ABB RAPID module: Weld1.mod

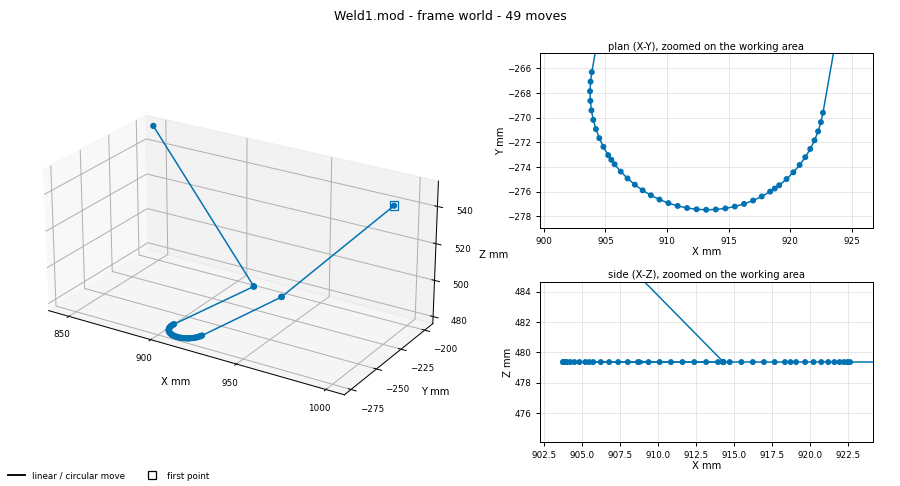
[picture p0: tool path of Weld1.mod in frame world, 49 of 50 moves have a stored position in this frame; points joined in program order, loops and branches not executed]
%%%
  VERSION:1
  LANGUAGE:ENGLISH
%%%
MODULE MOD_Weld1

    ! -------------------------------
    ! Define customized variables here
    ! ...

	! Tool variables:
	PERS tooldata Weldgun := [TRUE,[[-4.000,0.000,371.300],[0.92387953,0.00000000,0.38268343,0.00000001]],[1,[0,0,20],[1,0,0,0],0,0,0.005]];

	! Reference variables:
	PERS wobjdata WeldingReference := [FALSE, TRUE, "", [[0,0,0],[1,0,0,0]],[[907.213,-302.346,276.168],[0.70442562,0.70442562,-0.06151869,-0.06151869]]];

	PROC Main()
		ConfJ \On;
		ConfL \Off;
		! Program generated by VerticalBot Studio for ABB IRB 2600-12/1.65 on 25/10/2026 12:00:00
		! Using nominal kinematics.
		! show Weld gun
		MoveAbsJ [[-12.555800,6.650190,11.177100,0.026927,72.173900,-2.607590],[9E+09,9E+09,9E+09,9E+09,9E+09,9E+09]],v1000,z1,Weldgun \WObj:=WeldingReference;
		SetRPM 70.0;
		MoveL [[80.178,273.912,-94.776],[0.27080492,-0.27039115,-0.65336714,0.65319576],[-1,0,-1,0],[9E+09,9E+09,9E+09,9E+09,9E+09,9E+09]],[16.67,500,5000,1000],z1,Weldgun \WObj:=WeldingReference;
		MoveL [[9.468,203.201,-94.776],[0.27080492,-0.27039115,-0.65336714,0.65319576],[-1,0,-1,0],[9E+09,9E+09,9E+09,9E+09,9E+09,9E+09]],[16.67,500,5000,1000],z1,Weldgun \WObj:=WeldingReference;
		GunOn;
		MoveL [[9.468,203.201,-94.776],[0.27080492,-0.27039115,-0.65336714,0.65319576],[-1,0,-1,0],[9E+09,9E+09,9E+09,9E+09,9E+09,9E+09]],[16.67,500,5000,1000],z1,Weldgun \WObj:=WeldingReference;
		MoveL [[9.521,203.201,-94.770],[0.27059813,-0.27059797,-0.65328151,0.65328145],[-1,0,-1,0],[9E+09,9E+09,9E+09,9E+09,9E+09,9E+09]],[16.67,500,5000,1000],z1,Weldgun \WObj:=WeldingReference;
		MoveL [[9.521,203.201,-34.925],[0.26109596,-0.28004323,-0.64928868,0.65713689],[-1,-1,-1,0],[9E+09,9E+09,9E+09,9E+09,9E+09,9E+09]],[16.67,500,5000,1000],z1,Weldgun \WObj:=WeldingReference;
		MoveL [[9.489,203.201,-34.145],[0.23425026,-0.30675221,-0.65944853,0.64510273],[-1,-1,0,0],[9E+09,9E+09,9E+09,9E+09,9E+09,9E+09]],[16.67,500,5000,1000],z1,Weldgun \WObj:=WeldingReference;
		MoveL [[9.394,203.201,-33.370],[0.20701375,-0.33294335,-0.66849979,0.63198265],[-1,-1,0,0],[9E+09,9E+09,9E+09,9E+09,9E+09,9E+09]],[16.67,500,5000,1000],z1,Weldgun \WObj:=WeldingReference;
		MoveL [[9.235,203.201,-32.605],[0.17943264,-0.35858122,-0.67642029,0.61780177],[-1,-1,0,0],[9E+09,9E+09,9E+09,9E+09,9E+09,9E+09]],[16.67,500,5000,1000],z1,Weldgun \WObj:=WeldingReference;
		MoveL [[9.014,203.201,-31.857],[0.15154219,-0.38361099,-0.68321444,0.60257415],[-1,-1,0,0],[9E+09,9E+09,9E+09,9E+09,9E+09,9E+09]],[16.67,500,5000,1000],z1,Weldgun \WObj:=WeldingReference;
		MoveL [[8.732,203.201,-31.128],[0.12340353,-0.40798899,-0.68885701,0.58633828],[-1,-1,0,0],[9E+09,9E+09,9E+09,9E+09,9E+09,9E+09]],[16.67,500,5000,1000],z1,Weldgun \WObj:=WeldingReference;
		MoveL [[8.391,203.201,-30.426],[0.09505233,-0.43169103,-0.69333556,0.56911660],[-1,-1,0,0],[9E+09,9E+09,9E+09,9E+09,9E+09,9E+09]],[16.67,500,5000,1000],z1,Weldgun \WObj:=WeldingReference;
		MoveL [[7.994,203.201,-29.753],[0.06655006,-0.45466761,-0.69664493,0.55093947],[-1,-1,0,0],[9E+09,9E+09,9E+09,9E+09,9E+09,9E+09]],[16.67,500,5000,1000],z1,Weldgun \WObj:=WeldingReference;
		MoveL [[7.544,203.201,-29.116],[0.03792629,-0.47687790,-0.69878733,0.53183205],[-1,-1,0,0],[9E+09,9E+09,9E+09,9E+09,9E+09,9E+09]],[16.67,500,5000,1000],z1,Weldgun \WObj:=WeldingReference;
		MoveL [[7.042,203.201,-28.517],[0.01240330,-0.49395227,-0.70281556,0.51176909],[-1,-1,0,0],[9E+09,9E+09,9E+09,9E+09,9E+09,9E+09]],[16.67,500,5000,1000],z1,Weldgun \WObj:=WeldingReference;
		MoveL [[6.733,203.201,-28.192],[0.00416831,0.50587340,0.70291668,-0.49998286],[-1,-1,0,0],[9E+09,9E+09,9E+09,9E+09,9E+09,9E+09]],[16.67,500,5000,1000],z1,Weldgun \WObj:=WeldingReference;
		MoveL [[6.408,203.201,-27.883],[0.02374061,0.52184249,0.69941540,-0.48778571],[-1,-1,0,0],[9E+09,9E+09,9E+09,9E+09,9E+09,9E+09]],[16.67,500,5000,1000],z1,Weldgun \WObj:=WeldingReference;
		MoveL [[5.809,203.201,-27.381],[0.05240062,0.54140968,0.69785181,-0.46597487],[-1,-1,0,0],[9E+09,9E+09,9E+09,9E+09,9E+09,9E+09]],[16.67,500,5000,1000],z1,Weldgun \WObj:=WeldingReference;
		MoveL [[5.172,203.201,-26.930],[0.08097272,0.56005587,0.69511960,-0.44338425],[-1,-1,0,0],[9E+09,9E+09,9E+09,9E+09,9E+09,9E+09]],[16.67,500,5000,1000],z1,Weldgun \WObj:=WeldingReference;
		MoveL [[4.499,203.201,-26.534],[0.10940637,0.57776774,0.69121158,-0.42004909],[-1,-1,0,0],[9E+09,9E+09,9E+09,9E+09,9E+09,9E+09]],[16.67,500,5000,1000],z1,Weldgun \WObj:=WeldingReference;
		MoveL [[3.797,203.201,-26.193],[0.13765258,0.59450380,0.68614585,-0.39600615],[-1,-1,0,0],[9E+09,9E+09,9E+09,9E+09,9E+09,9E+09]],[16.67,500,5000,1000],z1,Weldgun \WObj:=WeldingReference;
		MoveL [[3.068,203.201,-25.912],[0.16567219,0.61024237,0.67992465,-0.37129428],[-1,-1,0,0],[9E+09,9E+09,9E+09,9E+09,9E+09,9E+09]],[16.67,500,5000,1000],z1,Weldgun \WObj:=WeldingReference;
		MoveL [[2.320,203.201,-25.690],[0.19341081,0.62495524,0.67255736,-0.34596213],[-1,-1,0,0],[9E+09,9E+09,9E+09,9E+09,9E+09,9E+09]],[16.67,500,5000,1000],z1,Weldgun \WObj:=WeldingReference;
		MoveL [[1.555,203.201,-25.531],[0.22082406,0.63861348,0.66406224,-0.32004826],[-1,-1,0,0],[9E+09,9E+09,9E+09,9E+09,9E+09,9E+09]],[16.67,500,5000,1000],z1,Weldgun \WObj:=WeldingReference;
		MoveL [[0.780,203.201,-25.436],[0.24786932,0.65119902,0.65444982,-0.29359169],[-1,-1,0,0],[9E+09,9E+09,9E+09,9E+09,9E+09,9E+09]],[16.67,500,5000,1000],z1,Weldgun \WObj:=WeldingReference;
		MoveL [[0.000,203.201,-25.404],[0.27449275,0.66268723,0.64373837,-0.26664635],[-1,-1,0,0],[9E+09,9E+09,9E+09,9E+09,9E+09,9E+09]],[16.67,500,5000,1000],z1,Weldgun \WObj:=WeldingReference;
		MoveL [[-0.780,203.201,-25.436],[0.30065949,0.67306272,0.63194229,-0.23924755],[-1,-1,0,0],[9E+09,9E+09,9E+09,9E+09,9E+09,9E+09]],[16.67,500,5000,1000],z1,Weldgun \WObj:=WeldingReference;
		MoveL [[-1.555,203.201,-25.531],[0.32631571,0.68230801,0.61908153,-0.21145189],[-1,0,1,0],[9E+09,9E+09,9E+09,9E+09,9E+09,9E+09]],[16.67,500,5000,1000],z1,Weldgun \WObj:=WeldingReference;
		MoveL [[-2.320,203.201,-25.690],[0.35142970,0.69040355,0.60518073,-0.18329319],[-1,0,1,0],[9E+09,9E+09,9E+09,9E+09,9E+09,9E+09]],[16.67,500,5000,1000],z1,Weldgun \WObj:=WeldingReference;
		MoveL [[-3.068,203.201,-25.912],[0.37594474,0.69734095,0.59026085,-0.15483308],[-1,0,1,0],[9E+09,9E+09,9E+09,9E+09,9E+09,9E+09]],[16.67,500,5000,1000],z1,Weldgun \WObj:=WeldingReference;
		MoveL [[-3.797,203.201,-26.193],[0.39983154,0.70309811,0.57435509,-0.12611111],[-1,0,1,0],[9E+09,9E+09,9E+09,9E+09,9E+09,9E+09]],[16.67,500,5000,1000],z1,Weldgun \WObj:=WeldingReference;
		MoveL [[-4.499,203.201,-26.534],[0.42304339,0.70768163,0.55747448,-0.09717615],[-1,0,1,0],[9E+09,9E+09,9E+09,9E+09,9E+09,9E+09]],[16.67,500,5000,1000],z1,Weldgun \WObj:=WeldingReference;
		MoveL [[-5.172,203.201,-26.930],[0.44554480,0.71107104,0.53966024,-0.06807809],[-1,0,1,0],[9E+09,9E+09,9E+09,9E+09,9E+09,9E+09]],[16.67,500,5000,1000],z1,Weldgun \WObj:=WeldingReference;
		MoveL [[-5.809,203.201,-27.381],[0.46730140,0.71326404,0.52093536,-0.03886082],[-1,0,1,0],[9E+09,9E+09,9E+09,9E+09,9E+09,9E+09]],[16.67,500,5000,1000],z1,Weldgun \WObj:=WeldingReference;
		MoveL [[-6.408,203.201,-27.883],[0.48819595,0.71113015,0.50576611,-0.01261974],[-1,0,1,0],[9E+09,9E+09,9E+09,9E+09,9E+09,9E+09]],[16.67,500,5000,1000],z1,Weldgun \WObj:=WeldingReference;
		MoveL [[-6.731,203.201,-28.191],[0.49992546,0.71126987,0.49411825,0.00410579],[-1,0,1,0],[9E+09,9E+09,9E+09,9E+09,9E+09,9E+09]],[16.67,500,5000,1000],z1,Weldgun \WObj:=WeldingReference;
		MoveL [[-7.042,203.201,-28.517],[0.51134749,0.71391546,0.47777457,0.02408169],[-1,0,1,0],[9E+09,9E+09,9E+09,9E+09,9E+09,9E+09]],[16.67,500,5000,1000],z1,Weldgun \WObj:=WeldingReference;
		MoveL [[-7.544,203.201,-29.116],[0.53050914,0.71232829,0.45640294,0.05333687],[-1,0,1,0],[9E+09,9E+09,9E+09,9E+09,9E+09,9E+09]],[16.67,500,5000,1000],z1,Weldgun \WObj:=WeldingReference;
		MoveL [[-7.994,203.201,-29.753],[0.54878026,0.70953905,0.43426730,0.08250137],[-1,0,1,0],[9E+09,9E+09,9E+09,9E+09,9E+09,9E+09]],[16.67,500,5000,1000],z1,Weldgun \WObj:=WeldingReference;
		MoveL [[-8.391,203.201,-30.426],[0.56612441,0.70556165,0.41139698,0.11152774],[-1,0,1,0],[9E+09,9E+09,9E+09,9E+09,9E+09,9E+09]],[16.67,500,5000,1000],z1,Weldgun \WObj:=WeldingReference;
		MoveL [[-8.732,203.201,-31.128],[0.58251728,0.70039316,0.38784300,0.14035973],[-1,0,1,0],[9E+09,9E+09,9E+09,9E+09,9E+09,9E+09]],[16.67,500,5000,1000],z1,Weldgun \WObj:=WeldingReference;
		MoveL [[-9.014,203.201,-31.857],[0.59792965,0.69404912,0.36363243,0.16895976],[-1,0,1,0],[9E+09,9E+09,9E+09,9E+09,9E+09,9E+09]],[16.67,500,5000,1000],z1,Weldgun \WObj:=WeldingReference;
		MoveL [[-9.235,203.201,-32.605],[0.61233261,0.68654186,0.33880881,0.19727554],[-1,0,1,0],[9E+09,9E+09,9E+09,9E+09,9E+09,9E+09]],[16.67,500,5000,1000],z1,Weldgun \WObj:=WeldingReference;
		MoveL [[-9.394,203.201,-33.370],[0.62571166,0.67787385,0.31341661,0.22525981],[-1,0,1,0],[9E+09,9E+09,9E+09,9E+09,9E+09,9E+09]],[16.67,500,5000,1000],z1,Weldgun \WObj:=WeldingReference;
		MoveL [[-9.489,203.201,-34.145],[0.63803534,0.66806855,0.28749564,0.25286671],[-1,0,1,0],[9E+09,9E+09,9E+09,9E+09,9E+09,9E+09]],[16.67,500,5000,1000],z1,Weldgun \WObj:=WeldingReference;
		MoveL [[-9.521,203.201,-34.925],[0.65328148,0.65328148,0.27059805,0.27059805],[-1,0,1,0],[9E+09,9E+09,9E+09,9E+09,9E+09,9E+09]],[16.67,500,5000,1000],z1,Weldgun \WObj:=WeldingReference;
		MoveL [[-9.521,203.201,-94.770],[0.65328148,0.65328148,0.27059805,0.27059805],[-1,0,1,0],[9E+09,9E+09,9E+09,9E+09,9E+09,9E+09]],[16.67,500,5000,1000],z1,Weldgun \WObj:=WeldingReference;
		MoveL [[-9.470,203.201,-94.776],[0.65328148,0.65328148,0.27059805,0.27059805],[-1,0,1,0],[9E+09,9E+09,9E+09,9E+09,9E+09,9E+09]],[16.67,500,5000,1000],z1,Weldgun \WObj:=WeldingReference;
		GunOff;
		MoveL [[-9.470,203.201,-94.776],[0.65328148,0.65328148,0.27059805,0.27059805],[-1,0,1,0],[9E+09,9E+09,9E+09,9E+09,9E+09,9E+09]],v1000,z1,Weldgun \WObj:=WeldingReference;
		MoveL [[-80.181,273.912,-94.776],[0.65328148,0.65328148,0.27059805,0.27059805],[-1,0,1,0],[9E+09,9E+09,9E+09,9E+09,9E+09,9E+09]],v1000,z1,Weldgun \WObj:=WeldingReference;
	ENDPROC

ENDMODULE
